Staubli VAL3: main.pgx

program main()
begin
  close(tCurrentTool)
  pPointRs.config.shoulder = lefty
  pPointRs2.config.shoulder = lefty
  mCurrentSpeed.tvel = 100.00
  mCurrentSpeed.blend = joint
  mCurrentSpeed.reach = 0.010
  mCurrentSpeed.leave = 0.010
  // Program ConfProg start
  // Program generated by RoboDK v6.0.7 for Staubli TP80 on XX/XX/XXXX 18:00:00
  // Using nominal kinematics.
  call MoveLine(-640.584,506.980,371.534,136.262,30.757,-130.375)
  pPointRs.config.shoulder = righty
  call MoveLine(-607.850,543.849,363.215,136.262,30.757,-130.375)
  pPointRs.config.shoulder = lefty
  call MoveLine(-602.951,596.788,316.595,136.262,30.757,-130.375)
  call MoveJoint(10.00000,20.00000,-30.00000,40.00000)
  call MoveJoint(-170.00000,45.00000,-45.00000,-170.00000)
  call MoveCirc(-353.026,-90.135,331.702,164.619,39.324,-168.579,-624.230,571.208,454.620,81.604,51.756,-128.588)

  waitEndMove()
  // Program ConfProg end

end
